Fanuc KAREL source: KA00041.KL

PROGRAM KA00041
%NOLOCKGROUP
VAR
  SRC: STRING[80]
  DST: POSITION
BEGIN
  SRC = 'A'
  DST = SRC
END KA00041
